Fanuc KAREL source: kd00012.KL

-- PROVISIONAL review KL for V1013-1; original PC SHA256 c984fb1331879fceb9ab58e585488cb6b41bced4ff5fe559da90ea0f08a58b18
-- Incomplete behavior may be omitted. Consult companion uncertainty JSON. Do not deploy.
PROGRAM KD00012
%NOLOCKGROUP
VAR
  I : INTEGER
  J : INTEGER
  B : BOOLEAN
  R : REAL
  S : STRING[80]
BEGIN
  -- UNRESOLVED_PC offsets 5-9; opcodes 9D,9D,1A
  -- UNRESOLVED_PC offsets 14-18; opcodes 7F
END KD00012
